(* Generated by scripts/make_testbench.py. Do not edit. *)
DATA_BLOCK "DB_TestResult"
{ S7_Optimized_Access := 'TRUE' }
VERSION : 0.1
NON_RETAIN
   VAR
      Done : Bool;
      CasesTotal : Int;
      CasesRun : Int;
      CasesPassed : Int;
      CasesFailed : Int;
      FirstFailedCase : Int;
      FirstFailedCheck : Int;
      CasePassed : Array[1..7] of Bool;
   END_VAR
BEGIN
END_DATA_BLOCK

DATA_BLOCK "TB_BENCH_DB"
{ S7_Optimized_Access := 'TRUE' }
VERSION : 0.1
NON_RETAIN
"TB_BENCH"
BEGIN
END_DATA_BLOCK
